(* IEC 61131-3 sources: SemantiST/compiler/intake/normalize/probes/elseif-keyword, 2 files *)

(* ---- original.st ---- *)
FUNCTION CLASSIFY : INT
VAR_INPUT
    A : INT;
END_VAR
IF A = 1 THEN
    CLASSIFY := 10;
ELSEIF A = 2 THEN
    CLASSIFY := 20;
ELSE
    CLASSIFY := 30;
END_IF;
END_FUNCTION

FUNCTION main : DINT
printf('%d %d %d$N', CLASSIFY(1), CLASSIFY(2), CLASSIFY(3));
main := 0;
END_FUNCTION

(* ---- rewritten.st ---- *)
FUNCTION CLASSIFY : INT
VAR_INPUT
    A : INT;
END_VAR
IF A = 1 THEN
    CLASSIFY := 10;
ELSIF A = 2 THEN
    CLASSIFY := 20;
ELSE
    CLASSIFY := 30;
END_IF;
END_FUNCTION

FUNCTION main : DINT
printf('%d %d %d$N', CLASSIFY(1), CLASSIFY(2), CLASSIFY(3));
main := 0;
END_FUNCTION
